// TIA Portal V20 export
// export: Created 2026-10-12T05:35:26.8814443Z, ExportSetting WithDefaults, DisplayName Totally Integrated Automation Portal, DisplayVersion V20, DisplayName TIA Portal Openness, DisplayVersion V20, DisplayName TIA Portal Teamcenter Gateway, DisplayVersion V20, DisplayName TIA Portal Version Control Interface, DisplayVersion V20, DisplayName SINAMICS Startdrive Advanced, DisplayVersion V20 SP1 Update 2, DisplayName SINAMICS Startdrive G110M, G120, G120C, G120D, G120P, G115D, DisplayVersion V20 SP1 Update 2, DisplayName SINAMICS Startdrive G130, G150, S120, S150, SINAMICS MV, G220, S200, S210, DisplayVersion V20 SP1 Update 2, DisplayName STEP 7 Professional, DisplayVersion V20, DisplayName STEP 7 Safety, DisplayVersion V20, DisplayName WinCC Basic/Comfort/Advanced, DisplayVersion V20, DisplayName WinCC Professional, DisplayVersion V20, DisplayName WinCC Unified, DisplayVersion V20
FUNCTION_BLOCK "FB_DeclarationCylinder"   // FB1, SCL
{ S7_Optimized_Access := 'TRUE' }
VERSION : 0.1
// Generated frame v0.11; change the declaration, then regenerate.
// stored: AutoNumber true, IsIECCheckEnabled false, IsRetainMemResEnabled false, MemoryReserve 100, SetENOAutomatically false, UDAEnableTagReadback false
   VAR_INPUT
      Execute { ExternalWritable := 'False'} : Bool;
      Abort { ExternalWritable := 'False'} : Bool;
      Command { ExternalWritable := 'False'} : DInt;
      ParCmd { ExternalWritable := 'False'} : "ST_DeclarationParCmd";
      ParentIndex { ExternalAccessible := 'False'; ExternalVisible := 'False'; ExternalWritable := 'False'} : DInt;
      Startup { ExternalAccessible := 'False'; ExternalVisible := 'False'; ExternalWritable := 'False'} : Bool;
   END_VAR
   VAR_OUTPUT
      Busy { ExternalWritable := 'False'} : Bool;
      Done { ExternalWritable := 'False'} : Bool;
      Error { ExternalWritable := 'False'} : Bool;
      Aborted { ExternalWritable := 'False'} : Bool;
      Held { ExternalWritable := 'False'} : Bool;
      ErrorID { ExternalWritable := 'False'} : DWord;
      Timing { ExternalWritable := 'False'} : "ST_ModuleTiming";
      OutCmd { ExternalWritable := 'False'} : "ST_DeclarationOutCmd";
      OutImm { ExternalWritable := 'False'} : "ST_DeclarationOutImm";
   END_VAR
   VAR_IN_OUT
      Hal : "ST_DeclarationLeafHal";
   END_VAR
   VAR
      Status { ExternalWritable := 'False'; S7_SetPoint := 'True'} : "ST_ModuleStatus";
      Core { ExternalAccessible := 'False'; ExternalVisible := 'False'; ExternalWritable := 'False'; S7_SetPoint := 'True'} : "FRK_Core";
      ParCfg { ExternalWritable := 'False'; S7_SetPoint := 'True'} : "ST_DeclarationParCfg";
      LatchedParCmd { ExternalAccessible := 'False'; ExternalVisible := 'False'; ExternalWritable := 'False'; S7_SetPoint := 'True'} : "ST_DeclarationParCmd";
      Device { ExternalAccessible := 'False'; ExternalVisible := 'False'; ExternalWritable := 'False'; S7_SetPoint := 'True'} : "ST_DeclarationOutImm";
      ConfigStageParCfg { ExternalAccessible := 'False'; ExternalVisible := 'False'; ExternalWritable := 'False'; S7_SetPoint := 'True'} : "ST_DeclarationParCfg";
      ConfigDefaultParCfg { ExternalAccessible := 'False'; ExternalVisible := 'False'; ExternalWritable := 'False'; S7_SetPoint := 'True'} : "ST_DeclarationParCfg";
      ConfigStaged { ExternalAccessible := 'False'; ExternalVisible := 'False'; ExternalWritable := 'False'} : Bool;
      Catalog { ExternalAccessible := 'False'; ExternalVisible := 'False'; ExternalWritable := 'False'; S7_SetPoint := 'True'} : Array[1..12] of "ST_CommandInfo";
      CatalogCount { ExternalAccessible := 'False'; ExternalVisible := 'False'; ExternalWritable := 'False'} : Int;
      ManConditions { ExternalAccessible := 'False'; ExternalVisible := 'False'; ExternalWritable := 'False'; S7_SetPoint := 'True'} : Array[1..16] of "FRK_ManualConditionRow";
      ManualOwned { ExternalAccessible := 'False'; ExternalVisible := 'False'; ExternalWritable := 'False'} : Bool;
   END_VAR
   VAR_TEMP
      InstancePath : WString[254];
   END_VAR
   VAR CONSTANT
      EXEC_READY : DInt := 0;
      MODULE_TIER : DInt := 3;
   END_VAR
BEGIN

   // ---- GENERATED: setup
   IF #Startup OR NOT #Core.Named THEN
       #InstancePath := GetInstancePath(size := 0);
       "FRK_SetIdentity"(Core := #Core,
                         Status := #Status,
                         InstancePath := #InstancePath,
                         ModuleType := 3,
                         TypeId := 3,
                         Capabilities := DWORD#16#00000000,
                         ParentIndex := #ParentIndex,
                         TypeKey := 'Fraktal.Declaration.Cylinder');
       #CatalogCount := 7;
       #Catalog[1].Value := 1;
       #Catalog[1].Label := 'Finish';
       #Catalog[1].Style := 0;
       #Catalog[2].Value := 2;
       #Catalog[2].Label := 'Wait';
       #Catalog[2].Style := 0;
       #Catalog[3].Value := 3;
       #Catalog[3].Label := 'Hold';
       #Catalog[3].Style := 0;
       #Catalog[4].Value := 4;
       #Catalog[4].Label := 'Fault';
       #Catalog[4].Style := 0;
       #Catalog[5].Value := 5;
       #Catalog[5].Label := 'Pending';
       #Catalog[5].Style := 0;
       #Catalog[6].Value := 6;
       #Catalog[6].Label := 'Instant';
       #Catalog[6].Style := 0;
       #Catalog[7].Value := 7;
       #Catalog[7].Label := 'Adopt';
       #Catalog[7].Style := 0;
   END_IF;
   IF #Startup THEN "FRK_CfgRestore_DeclarationCylinder"(Core := #Core,
                                                             Status := #Status,
                                                             ParCfg := #ParCfg,
                                                             ConfigStageParCfg := #ConfigStageParCfg,
                                                             ConfigDefaultParCfg := #ConfigDefaultParCfg);
   END_IF;
   // ---- GENERATED: begin
   "FRK_Begin"(Core := #Core,
               Status := #Status,
               Execute := #Execute,
               Abort := #Abort,
               Command := #Command);
   IF #Core.EvInit THEN
       // ---- AUTHORED: Init
       #Device.InitCount := #Device.InitCount + 1;
       // ---- GENERATED: reaction end
   END_IF;
   IF #Core.EvCommandStart THEN
       #LatchedParCmd := #ParCmd;
       CASE #Core.Command OF
           1:
               "FRK_Start"(Core := #Core,
                           Status := #Status,
                           Supported := TRUE,
                           Timeout := #ParCfg.Timeout,
                           Label := 'Finish');
           2:
               "FRK_Start"(Core := #Core,
                           Status := #Status,
                           Supported := TRUE,
                           Timeout := #ParCfg.Timeout,
                           Label := 'Wait');
           3:
               "FRK_Start"(Core := #Core,
                           Status := #Status,
                           Supported := TRUE,
                           Timeout := #ParCfg.Timeout,
                           Label := 'Hold');
           4:
               "FRK_Start"(Core := #Core,
                           Status := #Status,
                           Supported := TRUE,
                           Timeout := #ParCfg.Timeout,
                           Label := 'Fault');
           5:
               "FRK_Start"(Core := #Core,
                           Status := #Status,
                           Supported := TRUE,
                           Timeout := #ParCfg.Timeout,
                           Label := 'Pending');
           6:
               "FRK_Start"(Core := #Core,
                           Status := #Status,
                           Supported := TRUE,
                           Timeout := #ParCfg.Timeout,
                           Label := 'Instant');
           7:
               "FRK_Start"(Core := #Core,
                           Status := #Status,
                           Supported := TRUE,
                           Timeout := #ParCfg.Timeout,
                           Label := 'Adopt');
           ELSE
               "FRK_Start"(Core := #Core,
                           Status := #Status,
                           Supported := FALSE,
                           Timeout := T#0ms,
                           Label := '');
       END_CASE;
   END_IF;
   IF #Core.EvCommandStart THEN
       // ---- AUTHORED: CommandStart
       #Device.StartCount := #Device.StartCount + 1;
       #Device.Ordered := #Device.InitCount = 1;
       // ---- GENERATED: reaction end
   END_IF;
   // ---- AUTHORED: cyclic management
   #Device.CyclicCount := #Device.CyclicCount + 1;
   IF #Hal.BackgroundFault THEN
       "FRK_Fault"(Core := #Core,
                   Status := #Status,
                   ReasonCode := 2901,
                   Description := WSTRING#'test.background');
   END_IF;
   // ---- GENERATED: end management
   "FRK_RouteAbort"(Core := #Core,
                    Abort := #Abort);
   IF #Core.EvAbort THEN
       // ---- AUTHORED: Abort
       #Device.AbortCount := #Device.AbortCount + 1;
       // ---- GENERATED: reaction end
   END_IF;
   IF #Core.EvAbortInError THEN
       // ---- AUTHORED: AbortInError
       #Device.ErrorAbortCount := #Device.ErrorAbortCount + 1;
       // ---- GENERATED: reaction end
   END_IF;
   IF #Core.Dispatch AND #Core.RegIndex > 0 AND NOT "FRK_Registry".Fault THEN
       // ---- AUTHORED: dispatch
       #Device.DispatchCount := #Device.DispatchCount + 1;
       #Device.SeenValue := #LatchedParCmd.Value;
       CASE #Core.Command OF
           1:
               IF #Hal.Finish THEN
                   #OutCmd.Result := #LatchedParCmd.Value;
                   "FRK_Complete"(Core := #Core,
                                  Status := #Status);
               END_IF;
           2:
               #Device.SeenValue := #LatchedParCmd.Value;
           3:
               IF NOT #Hal.Permit THEN
                   "FRK_Hold"(Core := #Core,
                              Status := #Status,
                              ReasonCode := 2003,
                              Description := WSTRING#'test.permit');
               ELSIF #Hal.Finish THEN
                   "FRK_Complete"(Core := #Core,
                                  Status := #Status);
               END_IF;
           4:
               "FRK_Fault"(Core := #Core,
                           Status := #Status,
                           ReasonCode := 2901,
                           Description := WSTRING#'test.first');
               "FRK_Fault"(Core := #Core,
                           Status := #Status,
                           ReasonCode := 2001,
                           Description := WSTRING#'test.second');
           5:
               "FRK_Pending"(Core := #Core,
                             Status := #Status,
                             Diag := #Hal.Diag);
               "FRK_Pending"(Core := #Core,
                             Status := #Status,
                             Diag := #Hal.LaterDiag);
           6:
               "FRK_Complete"(Core := #Core,
                              Status := #Status);
           7:
               "FRK_AdoptFault"(Core := #Core,
                                Status := #Status,
                                Diag := #Hal.Diag);
           ELSE
               "FRK_Fault"(Core := #Core,
                           Status := #Status,
                           ReasonCode := 2008,
                           Description := WSTRING#'std.error.unsupportedHmiRequest');
       END_CASE;
       // ---- GENERATED: end dispatch
   END_IF;
   "FRK_End"(Core := #Core,
             Status := #Status,
             Busy => #Busy,
             Done => #Done,
             Error => #Error,
             Aborted => #Aborted,
             Held => #Held,
             ErrorID => #ErrorID,
             Timing => #Timing);
   // ---- AUTHORED: unconditional cyclic/derived data
   #Device.Sample := #Hal.Sample;
   #Device.Output := #Core.Exec = 1 AND NOT #Core.Held AND #Hal.Permit;
   #OutImm := #Device;
   // ---- GENERATED: frame end
END_FUNCTION_BLOCK
